// TIA Portal V20 export
TYPE "Keyence_IV3"
   STRUCT
      Status : Struct
         Warning_clear_request : Bool;   // Fordert das Löschen der Warnungen an
         Results_available : Bool;   // Ergebnisdaten sind verfügbar
         Result_update_complete : Bool;   // Durch einen Statuswechsel (0-1 oder 1-0) wird angegeben ob die Ergebnisdaten aktualisiert
         Busy : Bool;   // Während dieses Bit auf 1 ist, kann kein Trigger verarbeitet werden
         Imaging : Bool;   // Bildaufnahme wird ausgeführt
         RUN : Bool;   // Der Vision-Sensor ist im Run-Modus und es ist kein Systemfehler aufgetreten.
         Ready : Bool;   // Der Vision-Sensor ist komplett gestartet und betriebsbereit.
         Trigger_Ready : Bool;   // Dieses Bit wird ausgegeben, wenn der Trigger empfangen werden kann
         SD_card_Status : Bool;   // Dieses Bit wird ausgegeben, wenn die SD-Karte korrekt identifiziert wurde.
         SD_card_full : Bool;   // Dieses Bit wird ausgegeben, wenn der freie Speicherplatz auf der SD-Karte 100 MB oder weniger beträgt
         Warning : Bool;   // Warnung vorhanden
         Error_status : Bool;   // Fehler vorhanden
      END_STRUCT;
      Trigger : Struct
         Trigger_request : Bool;   // Fordert einen Trigger an
         Trigger_response : Bool;   // Speichert die Antwort des externen Triggers
         Overall_judgment_OK : Bool;   // Zeigt das Gesamtstatusergebnis an (OK)
         Busy : Bool;   // Während dieses Bit auf 1 ist, kann kein Trigger verarbeitet werden.
      END_STRUCT;
      Device_Result : Struct
         OveralljudgmentOK : Bool;   // Zeigt das Gesamtstatusergebnis an (OK)
         OveralljudgmentNG : Bool;   // Zeigt das Gesamtstatusergebnis an (NG)
         Positionscorrection : Bool;   // Ergebnis der Positionskorrektur
         Tool : Array[1..16] of Bool;   // Zeigt das Ergebnis von Werkzeug X an
      END_STRUCT;
      ToolX_Result : Struct
         Tool_Number : Int;   // Nummer des Werkzeugs, welches abgefragt werden soll
         Error : Bool;   // Gibt an, ob die Werkzeugnummer gültig ist
         Tool_matchingrate_max : Bool;   // Maximaler Übereinstimmungsgrad für Werkzeug
         Tool_matchingrate_min : Bool;   // Minimaler Übereinstimmungsgrad für Werkzeug
         Tool_lower_threshold : Bool;   // Unterer Grenzwert des Übereinstimmungsgrads für Werkzeug
         Tool_upper_threshold : Bool;   // Oberer Grenzwert des Übereinstimmungsgrads für Werkzeug
      END_STRUCT;
      Programm_Change : Struct
         SwitchProgram : Bool;   // Fordert einen Programmwechsel an
         ProgramNumber : UInt;   // Angabe der Programmnummer für einen Programmwechsel
         CurrentProgram : UInt;   // Aktuelle Programmnummer
         Programswitchresponse : Bool;   // Speichert die Programmwechselantwort
         Programswitchingfailed : Bool;   // Dieses Bit wird aktiviert, wenn der Trigger fehlgeschlagen ist
      END_STRUCT;
   END_STRUCT;
END_TYPE
